(*
SPDX-FileCopyrightText: © 2026 Oleksandr Tiutyk <trofimich@gmail.com>
SPDX-License-Identifier: MIT
License: https://opensource.org/license/mit
*)

(*!
<summary>
Beckhoff strain gauge / resistor bridge output control channel process image.
</summary>
<description>
Encapsulates a 16-bit control word for calibration, tare, and filtering commands on measuring bridge terminals
(e.g. EL3356).
When used for I/O, link located fields or their containing buffers to the matching selected PDOs.
The record is not a packed wire buffer; compiler padding is not part of the device specification.
Unlinked/default values do not prove valid I/O. The caller evaluates bus/channel validity before use.
Use one owner task per instance and externally synchronize other access; multi-field snapshots are not atomic.
Copies store data without creating hardware links. Keep borrowed field references valid while consumers are bound.
This passive record performs no validation, synchronization, configuration or protocol advancement.
</description>
*)
TYPE STRAIN_GAUGE_OUTPUT_CHANNEL :
STRUCT
	Control AT %Q* : WORD;
END_STRUCT
END_TYPE

(* stored: Version 1.1.0.1, ProductVersion 3.1.4026.20
   DUT STRAIN_GAUGE_OUTPUT_CHANNEL: Id {3146ac6b-a9fc-4681-a757-3b6321b88d3e} *)
